// TIA Portal V20 export
// export: Created 2026-10-21T10:56:20.5683147Z, ExportSetting None, DisplayName Totally Integrated Automation Portal, DisplayVersion V20, DisplayName TIA Portal Openness, DisplayVersion V20, DisplayName TIA Portal Version Control Interface, DisplayVersion V20, DisplayName STEP 7 Professional, DisplayVersion V20, DisplayName STEP 7 Safety, DisplayVersion V20, DisplayName WinCC Basic/Comfort/Advanced, DisplayVersion V20, DisplayName WinCC Unified, DisplayVersion V20
ORGANIZATION_BLOCK "Main"   // OB1, SCL, ProgramCycle
{ S7_Optimized_Access := 'TRUE' }
// stored: SetENOAutomatically false
   VAR_INPUT
      Initial_Call : Bool;   // Initial call of this OB
      Remanence : Bool;   // =True, if remanent data are available
   END_VAR
BEGIN

   // Arnes de prueba para FC_Escalado (bloques-de-funcion/fc-escalado/arnes-ob1.md).
   //
   // Las seis variables de test son REAL: la API de PLCSIM Advanced resuelve y escribe
   // simbolos REAL de forma nativa, mientras que el bloque recibe INT. El arnes hace la
   // conversion con REAL_TO_INT, que trunca hacia cero, y los valores de prueba se
   // mantienen dentro del rango INT.
   //
   // Mapa de tags (tabla Agent_Escalado):
   //   RawValue    entrada  valor crudo de la entrada analogica
   //   RawMin      entrada  raw del minimo de escala
   //   RawMax      entrada  raw del maximo de escala
   //   ScaleMin    entrada  valor de ingenieria del raw minimo
   //   ScaleMax    entrada  valor de ingenieria del raw maximo
   //   ScaledValue salida   valor escalado
   "FC_Escalado"(iValorCrudo := REAL_TO_INT("RawValue"),
                 iRawMin := REAL_TO_INT("RawMin"),
                 iRawMax := REAL_TO_INT("RawMax"),
                 rEscalaMin := "ScaleMin",
                 rEscalaMax := "ScaleMax",
                 rEscalado => "ScaledValue");
END_ORGANIZATION_BLOCK
